TYPE ST_PatchProcessSettings :
STRUCT
    lrDriveMotorVelocity : LREAL := 40.0;
    lrPatchFeedRollVelocity : LREAL := 200.0;
    lrWasteRollVelocity : LREAL := 50.0;
    udiReleaseMs : UDINT := 5000;
    udiAirBlowDelayMs : UDINT := 1500;
    // M1 run-on after the left optical clears; milliseconds.
    udiDriveStopDelayMs : UDINT := 2000;
END_STRUCT
END_TYPE

(* stored: Version 1.1.0.1, ProductVersion 3.1.4026.18
   DUT ST_PatchProcessSettings: Id {122c61c9-499d-42ab-af1a-dfbd125f9c0c} *)
